Fanuc KAREL source: KB00191.KL

PROGRAM KB00191
%NOLOCKGROUP
%ENVIRONMENT TRANS
VAR
  P1: STRING[80]
  P2: BOOLEAN
  P3: INTEGER
BEGIN
  P1 = 'A'
  P2 = TRUE
  P3 = 1
  TRANSLATE(P1, P2, P3)
END KB00191
